(* PLC project FM_XJV1.project, Xinje company XS Studio V2.3.2a XS Studio V2.3.2a *)
(* stored: creationDateTime 2026-10-30T20:27:28.6587941, modificationDateTime 2026-10-30T00:07:23.1916909 *)

CONFIGURATION Application
  RESOURCE Application ON PLC
    TASK EtherCAT_Task(INTERVAL := T#4ms, PRIORITY := 1);
    PROGRAM PLC_PRG WITH EtherCAT_Task : PLC_PRG;
  END_RESOURCE
END_CONFIGURATION
